// TIA Portal V15.1 export
// export: Created 2026-11-02T18:55:11.2894745Z, ExportSetting WithDefaults, DisplayName Totally Integrated Automation Portal, DisplayVersion V15.1, DisplayName TIA Portal Openness, DisplayVersion V15.1, DisplayName STEP 7 Professional, DisplayVersion V15.1, DisplayName WinCC Professional, DisplayVersion V15.1
FUNCTION "Outputs" : Void   // FC2, LAD
TITLE = Outputs
{ S7_Optimized_Access := 'TRUE' }
VERSION : 0.1
// The only block that writes %Q (decisions/0006 rule 3)
// stored: AutoNumber false, IsIECCheckEnabled false, SetENOAutomatically False, UDAEnableTagReadback false
BEGIN

REGION Network 1: E1 — BR01 heat request TL (R1, H1)
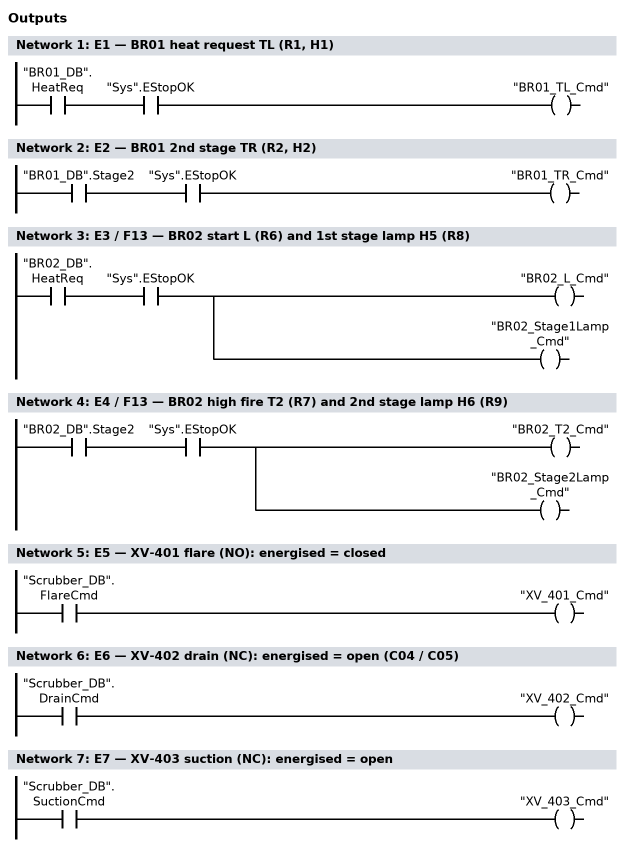
   RUNG wire#powerrail
      Contact( "BR01_DB".HeatReq )
      Contact( "Sys".EStopOK )
      Coil( "BR01_TL_Cmd" )
   END_RUNG
   // the same network as SCL:
   "BR01_TL_Cmd" := "BR01_DB".HeatReq AND "Sys".EStopOK;
END_REGION

REGION Network 2: E2 — BR01 2nd stage TR (R2, H2)
   RUNG wire#powerrail
      Contact( "BR01_DB".Stage2 )
      Contact( "Sys".EStopOK )
      Coil( "BR01_TR_Cmd" )
   END_RUNG
   // the same network as SCL:
   "BR01_TR_Cmd" := "BR01_DB".Stage2 AND "Sys".EStopOK;
END_REGION

REGION Network 3: E3 / F13 — BR02 start L (R6) and 1st stage lamp H5 (R8)
   RUNG wire#powerrail
      Contact( "BR02_DB".HeatReq )
      Contact( "Sys".EStopOK )
      wire#w1
      Coil( "BR02_L_Cmd" )
   END_RUNG
   RUNG wire#w1
      Coil( "BR02_Stage1Lamp_Cmd" )
   END_RUNG
   // the same network as SCL:
   "BR02_L_Cmd" := "BR02_DB".HeatReq AND "Sys".EStopOK;
   "BR02_Stage1Lamp_Cmd" := "BR02_L_Cmd";
END_REGION

REGION Network 4: E4 / F13 — BR02 high fire T2 (R7) and 2nd stage lamp H6 (R9)
   RUNG wire#powerrail
      Contact( "BR02_DB".Stage2 )
      Contact( "Sys".EStopOK )
      wire#w1
      Coil( "BR02_T2_Cmd" )
   END_RUNG
   RUNG wire#w1
      Coil( "BR02_Stage2Lamp_Cmd" )
   END_RUNG
   // the same network as SCL:
   "BR02_T2_Cmd" := "BR02_DB".Stage2 AND "Sys".EStopOK;
   "BR02_Stage2Lamp_Cmd" := "BR02_T2_Cmd";
END_REGION

REGION Network 5: E5 — XV-401 flare (NO): energised = closed
   RUNG wire#powerrail
      Contact( "Scrubber_DB".FlareCmd )
      Coil( "XV_401_Cmd" )
   END_RUNG
   // the same network as SCL:
   "XV_401_Cmd" := "Scrubber_DB".FlareCmd;
END_REGION

REGION Network 6: E6 — XV-402 drain (NC): energised = open (C04 / C05)
   RUNG wire#powerrail
      Contact( "Scrubber_DB".DrainCmd )
      Coil( "XV_402_Cmd" )
   END_RUNG
   // the same network as SCL:
   "XV_402_Cmd" := "Scrubber_DB".DrainCmd;
END_REGION

REGION Network 7: E7 — XV-403 suction (NC): energised = open
   RUNG wire#powerrail
      Contact( "Scrubber_DB".SuctionCmd )
      Coil( "XV_403_Cmd" )
   END_RUNG
   // the same network as SCL:
   "XV_403_Cmd" := "Scrubber_DB".SuctionCmd;
END_REGION
END_FUNCTION
